(* IEC 61131-3 sources: plc-process-lib/tests/POUs/Suites/FB_Util_Test, 29 files *)

(* ---- IsFiniteAboveSaneMaxReturnsFalse.method.decl.st ---- *)
// F_IsFinite: |x| > REAL_SANE_MAX — мусор (перепутан порядок слов Modbus): 1e31, -1e31 и
// наибольшее REAL — FALSE.
METHOD PRIVATE IsFiniteAboveSaneMaxReturnsFalse
VAR
    uBits : U_RealBits;      // значение REAL по битам IEEE 754
END_VAR

(* ---- IsFiniteInfReturnsFalse.method.decl.st ---- *)
// F_IsFinite: +Inf и -Inf — FALSE.
METHOD PRIVATE IsFiniteInfReturnsFalse
VAR
    uBits : U_RealBits;      // значение REAL по битам IEEE 754
END_VAR

(* ---- IsFiniteNaNReturnsFalse.method.decl.st ---- *)
// F_IsFinite: тихий NaN с обоими знаками и с полной мантиссой — FALSE (проверка R4 контракта).
METHOD PRIVATE IsFiniteNaNReturnsFalse
VAR
    uBits : U_RealBits;      // значение REAL по битам IEEE 754
END_VAR

(* ---- IsFiniteNormalReturnsTrue.method.decl.st ---- *)
// F_IsFinite: обычные числа, 0, -0, наименьшее денормализованное и граница ±REAL_SANE_MAX
// (включительно) — TRUE.
METHOD PRIVATE IsFiniteNormalReturnsTrue
VAR
    uBits : U_RealBits;      // значение REAL по битам IEEE 754
END_VAR

(* ---- LimitMonitorDisabledNeverSets.method.decl.st ---- *)
// Выключенная уставка (xEnable = FALSE) не взводит флаг: 10 с значение далеко за уставкой.
METHOD PRIVATE LimitMonitorDisabledNeverSets
VAR
    fbTime   : FB_FakeTime;       // подменное время
    fbLim    : FB_LimitMonitor;   // ФБ под тестом
    stLimCfg : ST_AiLimitCfg;     // параметры уставки
    iStep : INT;             // шаг цикла
    xEverSet : BOOL;            // флаг взводился хотя бы раз
END_VAR

(* ---- LimitMonitorDisabledNeverSets.method.impl.st ---- *)
coUnit.TEST('Util_LimitMonitor_Disabled_NeverSets');

stLimCfg.xEnable := FALSE;
stLimCfg.rSetpoint_eu := 50.0;
FOR iStep := 1 TO 100 DO
    fbTime.Advance(tStep := T#100MS);
    fbLim(rValue_eu := 90.0, xHighLimit := TRUE, stCfg := stLimCfg, itfTime := fbTime);
    xEverSet := xEverSet OR fbLim.xOut OR fbLim.xRaw;
END_FOR
AssertFalse(Condition := xEverSet, Message := 'disabled limit must never set the flag');

coUnit.TEST_FINISHED();

(* ---- LimitMonitorForceOffClearsImmediately.method.decl.st ---- *)
// xForceOff снимает флаг и сырой флаг в том же вызове, несмотря на задержку снятия 10 с; после
// снятия xForceOff флаг возвращается (значение по-прежнему выше уставки, задержки включения нет).
METHOD PRIVATE LimitMonitorForceOffClearsImmediately
VAR
    fbTime   : FB_FakeTime;       // подменное время
    fbLim    : FB_LimitMonitor;   // ФБ под тестом
    stLimCfg : ST_AiLimitCfg;     // параметры уставки
END_VAR

(* ---- LimitMonitorHighHysteresisClearsBelowSpMinusHyst.method.decl.st ---- *)
// Верхняя уставка 80, гистерезис 5: флаг при значении >= 80 (включительно), держится до 75
// включительно, снимается ниже 75; в зоне гистерезиса снятый флаг не возвращается.
METHOD PRIVATE LimitMonitorHighHysteresisClearsBelowSpMinusHyst
VAR
    fbTime   : FB_FakeTime;       // подменное время
    fbLim    : FB_LimitMonitor;   // ФБ под тестом
    stLimCfg : ST_AiLimitCfg;     // параметры уставки
END_VAR

(* ---- LimitMonitorLowHysteresisClearsAboveSpPlusHyst.method.decl.st ---- *)
// Нижняя уставка 20, гистерезис 2 — зеркально: флаг при значении <= 20, держится до 22
// включительно, снимается выше 22.
METHOD PRIVATE LimitMonitorLowHysteresisClearsAboveSpPlusHyst
VAR
    fbTime   : FB_FakeTime;       // подменное время
    fbLim    : FB_LimitMonitor;   // ФБ под тестом
    stLimCfg : ST_AiLimitCfg;     // параметры уставки
END_VAR

(* ---- LimitMonitorNonFiniteValueKeepsState.method.decl.st ---- *)
// Неконечное значение (NaN, ±Inf, больше REAL_SANE_MAX) флаг не меняет: -Inf не снимает
// взведённый флаг верхней уставки, +Inf не взводит снятый.
METHOD PRIVATE LimitMonitorNonFiniteValueKeepsState
VAR
    fbTime   : FB_FakeTime;       // подменное время
    fbLim    : FB_LimitMonitor;   // ФБ под тестом
    stLimCfg : ST_AiLimitCfg;     // параметры уставки
    uBits : U_RealBits;      // значение REAL по битам IEEE 754
END_VAR

(* ---- LimitMonitorOffDelayHoldsFlag.method.decl.st ---- *)
// Задержка снятия 2 с: сырой флаг снимается сразу, выходной держится до t0 + 1,9 с и снимается
// ровно в t0 + 2,0 с.
METHOD PRIVATE LimitMonitorOffDelayHoldsFlag
VAR
    fbTime   : FB_FakeTime;       // подменное время
    fbLim    : FB_LimitMonitor;   // ФБ под тестом
    stLimCfg : ST_AiLimitCfg;     // параметры уставки
    iStep : INT;             // шаг цикла
END_VAR

(* ---- LimitMonitorOffDelayHoldsFlag.method.impl.st ---- *)
coUnit.TEST('Util_LimitMonitor_OffDelay_HoldsFlag');

stLimCfg.xEnable := TRUE;
stLimCfg.rSetpoint_eu := 80.0;
stLimCfg.rHyst_eu := 2.0;
stLimCfg.tOffDelay := T#2S;
fbLim(rValue_eu := 85.0, xHighLimit := TRUE, stCfg := stLimCfg, itfTime := fbTime);
AssertTrue(Condition := fbLim.xOut, Message := 'flag set without on-delay');
fbLim(rValue_eu := 70.0, xHighLimit := TRUE, stCfg := stLimCfg, itfTime := fbTime);    // t0
AssertFalse(Condition := fbLim.xRaw, Message := 'raw flag cleared at once');
FOR iStep := 1 TO 19 DO
    fbTime.Advance(tStep := T#100MS);
    fbLim(rValue_eu := 70.0, xHighLimit := TRUE, stCfg := stLimCfg, itfTime := fbTime);
END_FOR
AssertTrue(Condition := fbLim.xOut, Message := 'flag held at t0 + 1.9 s');
fbTime.Advance(tStep := T#100MS);
fbLim(rValue_eu := 70.0, xHighLimit := TRUE, stCfg := stLimCfg, itfTime := fbTime);
AssertFalse(Condition := fbLim.xOut, Message := 'flag cleared exactly at t0 + 2.0 s');

coUnit.TEST_FINISHED();

(* ---- LimitMonitorOnDelayShortExcursionIgnored.method.decl.st ---- *)
// Задержка срабатывания 3 с: выброс 2,9 с за уставку флаг не взводит (сырой флаг — да);
// устойчивое превышение — флаг ровно через 3 с.
METHOD PRIVATE LimitMonitorOnDelayShortExcursionIgnored
VAR
    fbTime   : FB_FakeTime;       // подменное время
    fbLim    : FB_LimitMonitor;   // ФБ под тестом
    stLimCfg : ST_AiLimitCfg;     // параметры уставки
    iStep : INT;             // шаг цикла
    xEverSet : BOOL;            // флаг взводился хотя бы раз
END_VAR

(* ---- LimitMonitorOnDelayShortExcursionIgnored.method.impl.st ---- *)
coUnit.TEST('Util_LimitMonitor_OnDelay_ShortExcursionIgnored');

stLimCfg.xEnable := TRUE;
stLimCfg.rSetpoint_eu := 80.0;
stLimCfg.rHyst_eu := 2.0;
stLimCfg.tOnDelay := T#3S;
fbLim(rValue_eu := 85.0, xHighLimit := TRUE, stCfg := stLimCfg, itfTime := fbTime);    // t0
FOR iStep := 1 TO 29 DO                                                               // t0 + 2,9 с
    fbTime.Advance(tStep := T#100MS);
    fbLim(rValue_eu := 85.0, xHighLimit := TRUE, stCfg := stLimCfg, itfTime := fbTime);
    xEverSet := xEverSet OR fbLim.xOut;
END_FOR
AssertTrue(Condition := fbLim.xRaw, Message := 'raw flag is set before the delay');
fbTime.Advance(tStep := T#100MS);
fbLim(rValue_eu := 70.0, xHighLimit := TRUE, stCfg := stLimCfg, itfTime := fbTime);    // t0 + 3,0 с
xEverSet := xEverSet OR fbLim.xOut;
AssertFalse(Condition := xEverSet, Message := 'excursion shorter than the on-delay must be ignored');
fbLim(rValue_eu := 85.0, xHighLimit := TRUE, stCfg := stLimCfg, itfTime := fbTime);    // t1
FOR iStep := 1 TO 29 DO
    fbTime.Advance(tStep := T#100MS);
    fbLim(rValue_eu := 85.0, xHighLimit := TRUE, stCfg := stLimCfg, itfTime := fbTime);
END_FOR
AssertFalse(Condition := fbLim.xOut, Message := 'no flag at t1 + 2.9 s');
fbTime.Advance(tStep := T#100MS);
fbLim(rValue_eu := 85.0, xHighLimit := TRUE, stCfg := stLimCfg, itfTime := fbTime);    // t1 + 3,0 с
AssertTrue(Condition := fbLim.xOut, Message := 'flag exactly at t1 + 3.0 s');

coUnit.TEST_FINISHED();

(* ---- LimitMonitorReenabledRestartsOnDelay.method.decl.st ---- *)
// Выключение уставки во время задержки срабатывания (2 с) сбрасывает отсчёт: после повторного
// включения в t0 + 1,6 с флаг — ровно через 2 с от включения, а не в t0 + 2,0 с.
METHOD PRIVATE LimitMonitorReenabledRestartsOnDelay
VAR
    fbTime   : FB_FakeTime;       // подменное время
    fbLim    : FB_LimitMonitor;   // ФБ под тестом
    stLimCfg : ST_AiLimitCfg;     // параметры уставки
    iStep : INT;             // шаг цикла
END_VAR

(* ---- LimitMonitorReenabledRestartsOnDelay.method.impl.st ---- *)
coUnit.TEST('Util_LimitMonitor_Reenabled_RestartsOnDelay');

stLimCfg.xEnable := TRUE;
stLimCfg.rSetpoint_eu := 80.0;
stLimCfg.tOnDelay := T#2S;
fbLim(rValue_eu := 90.0, xHighLimit := TRUE, stCfg := stLimCfg, itfTime := fbTime);    // t0
FOR iStep := 1 TO 15 DO                                                               // t0 + 1,5 с
    fbTime.Advance(tStep := T#100MS);
    fbLim(rValue_eu := 90.0, xHighLimit := TRUE, stCfg := stLimCfg, itfTime := fbTime);
END_FOR
stLimCfg.xEnable := FALSE;
fbLim(rValue_eu := 90.0, xHighLimit := TRUE, stCfg := stLimCfg, itfTime := fbTime);
AssertFalse(Condition := fbLim.xOut OR fbLim.xRaw, Message := 'disabled: flags cleared');
stLimCfg.xEnable := TRUE;
FOR iStep := 1 TO 5 DO                                                                // t0 + 1,6 … 2,0 с
    fbTime.Advance(tStep := T#100MS);
    fbLim(rValue_eu := 90.0, xHighLimit := TRUE, stCfg := stLimCfg, itfTime := fbTime);
END_FOR
AssertFalse(Condition := fbLim.xOut, Message := 'old timing must not complete after re-enable');
FOR iStep := 1 TO 15 DO                                                               // t0 + 3,5 с
    fbTime.Advance(tStep := T#100MS);
    fbLim(rValue_eu := 90.0, xHighLimit := TRUE, stCfg := stLimCfg, itfTime := fbTime);
END_FOR
AssertFalse(Condition := fbLim.xOut, Message := 'no flag 1.9 s after re-enable');
fbTime.Advance(tStep := T#100MS);
fbLim(rValue_eu := 90.0, xHighLimit := TRUE, stCfg := stLimCfg, itfTime := fbTime);    // t0 + 3,6 с
AssertTrue(Condition := fbLim.xOut, Message := 'flag 2.0 s after re-enable');

coUnit.TEST_FINISHED();

(* ---- RateLimitLrNonFiniteTargetOrZeroDtHoldsCurrent.method.decl.st ---- *)
// F_RateLimitLr: цель NaN (мусор Modbus) или шаг времени 0 — значение не меняется; скорость 0 — сразу к цели;
// текущее значение NaN — сразу к цели (как F_RateLimit, F-11).
METHOD PRIVATE RateLimitLrNonFiniteTargetOrZeroDtHoldsCurrent
VAR
    uBits : U_RealBits;      // значение REAL по битам IEEE 754
    lrOut : LREAL;           // результат F_RateLimitLr
    lrNaN : LREAL;           // NaN в LREAL
END_VAR

(* ---- RateLimitLrSmallStepNotLost.method.decl.st ---- *)
// F_RateLimitLr: состояние в LREAL — 1000 шагов по 1 мс со скоростью 0,003 ед./с от 70,0 дают 70,003 (в REAL
// приращение 3·10⁻⁶ меньше половины шага REAL рядом с 70 и терялось бы); спад — так же; цель достигается точно.
METHOD PRIVATE RateLimitLrSmallStepNotLost
VAR
    lrUp   : LREAL;          // рост: состояние рампы
    lrDown : LREAL;          // спад: состояние рампы
    iStep  : INT;            // шаг цикла
END_VAR

(* ---- RateLimitLrSmallStepNotLost.method.impl.st ---- *)
coUnit.TEST('Util_RateLimitLr_SmallStep_NotLost');

lrUp := 70.0;
lrDown := 70.0;
FOR iStep := 1 TO 1000 DO
    lrUp := F_RateLimitLr(lrCurrent := lrUp, rTarget := 100.0, rRateUp_ups := 0.003, rRateDown_ups := 0.003,
                          lrDt_s := 0.001);
    lrDown := F_RateLimitLr(lrCurrent := lrDown, rTarget := 0.0, rRateUp_ups := 0.003, rRateDown_ups := 0.003,
                            lrDt_s := 0.001);
END_FOR
// ожидаемое: 70 ± 0,003 · 1 с; допуск — шаг REAL скорости 0,003 · 1000 шагов
AssertEquals_LREAL(Expected := LREAL#70.003, Actual := lrUp, Delta := LREAL#1.0E-7, Message := 'ramp up not lost');
AssertEquals_LREAL(Expected := LREAL#69.997, Actual := lrDown, Delta := LREAL#1.0E-7, Message := 'ramp down not lost');
AssertEquals_LREAL(Expected := LREAL#42.5, Actual := F_RateLimitLr(lrCurrent := LREAL#42.49, rTarget := 42.5,
                   rRateUp_ups := 1.0, rRateDown_ups := 1.0, lrDt_s := 1.0), Delta := LREAL#0.0,
                   Message := 'reaches the target exactly');

coUnit.TEST_FINISHED();

(* ---- RateLimitNonFiniteCurrentJumpsToTarget.method.decl.st ---- *)
// F_RateLimit: текущее значение NaN (мусор прошлого шага) заменяется конечной целью — ограничитель
// не застревает на NaN.
METHOD PRIVATE RateLimitNonFiniteCurrentJumpsToTarget
VAR
    uBits : U_RealBits;      // значение REAL по битам IEEE 754
    rOut  : REAL;            // результат F_RateLimit
END_VAR

(* ---- RateLimitNonFiniteTargetHoldsCurrent.method.decl.st ---- *)
// F_RateLimit: цель NaN, +Inf или больше REAL_SANE_MAX (мусор из Modbus/ПИД) — значение удерживается.
METHOD PRIVATE RateLimitNonFiniteTargetHoldsCurrent
VAR
    uBits : U_RealBits;      // значение REAL по битам IEEE 754
    rOut  : REAL;            // результат F_RateLimit
END_VAR

(* ---- StartsWindowClearEmpties.method.decl.st ---- *)
// Clear очищает окно: пусков 0, освобождать нечего.
METHOD PRIVATE StartsWindowClearEmpties
VAR
    fbWin : FB_StartsWindow; // ФБ под тестом
END_VAR

(* ---- StartsWindowCountsOnlyLastHour.method.decl.st ---- *)
// FB_StartsWindow: пуски в 1:00, 1:20, 1:40 — в окне последнего часа их 3, 2, 1, 0 по мере
// старения. Источник: tools/reference/common.py, сценарий starts_window.
METHOD PRIVATE StartsWindowCountsOnlyLastHour
VAR
    fbWin : FB_StartsWindow; // ФБ под тестом
END_VAR

(* ---- StartsWindowExactlyOneHourOldNotCounted.method.decl.st ---- *)
// Граница окна: отметка ровно часовой давности уже не считается (ltNow - t < STARTS_WINDOW).
METHOD PRIVATE StartsWindowExactlyOneHourOldNotCounted
VAR
    fbWin : FB_StartsWindow; // ФБ под тестом
END_VAR

(* ---- StartsWindowRingCapacityMatchesConst.method.decl.st ---- *)
// Ёмкость кольца altStart равна GVL_Const.STARTS_WINDOW_MAX: индексы кольца считаются по константе,
// тест ловит расхождение, если границу массива запишут числом.
// Тест обращается к внутренней переменной ФБ намеренно: это проверка раскладки, а не API.
METHOD PRIVATE StartsWindowRingCapacityMatchesConst
VAR
    fbWin : FB_StartsWindow; // ФБ под тестом
    ltOne : LTIME;           // один элемент кольца
END_VAR

(* ---- StartsWindowRingFullOverwritesOldest.method.decl.st ---- *)
// Кольцо на STARTS_WINDOW_MAX = 30: 31 пуск с шагом 1 мин (1:00…1:30) — остаются 30 последних;
// в 1:30 при лимите 30 окно освободится через 31 мин (самый старый оставшийся — 1:01).
// Источник: tools/reference/common.py, сценарий starts_window.
METHOD PRIVATE StartsWindowRingFullOverwritesOldest
VAR
    fbWin : FB_StartsWindow; // ФБ под тестом
    ltStart : LTIME := LTIME#1H;   // время очередного пуска
    iStep : INT;             // шаг цикла
END_VAR

(* ---- StartsWindowRingFullOverwritesOldest.method.impl.st ---- *)
coUnit.TEST('Util_StartsWindow_RingFull_OverwritesOldest');

FOR iStep := 0 TO 30 DO
    fbWin.Register(ltNow := ltStart);
    ltStart := ltStart + LTIME#1M;
END_FOR
AssertEquals_UINT(Expected := 30, Actual := fbWin.Count(ltNow := LTIME#1H30M), Message := 'ring keeps 30 starts');
AssertEquals_LTIME(Expected := LTIME#31M, Actual := fbWin.TimeToFree(ltNow := LTIME#1H30M, uiMax := 30),
                   Message := 'the start of 1:00 was overwritten, the oldest kept is 1:01');

coUnit.TEST_FINISHED();

(* ---- StartsWindowTimeBackwardsDropsFutureStamps.method.decl.st ---- *)
// Время назад: отметки «из будущего» удаляются и в Count, и в Register; окно остаётся упорядоченным.
METHOD PRIVATE StartsWindowTimeBackwardsDropsFutureStamps
VAR
    fbWin : FB_StartsWindow; // ФБ под тестом
END_VAR

(* ---- StartsWindowTimeToFreeReportsRemaining.method.decl.st ---- *)
// TimeToFree: пуски 1:00, 1:10, 1:20; в 1:30 при лимите 3 — 30 мин, при лимите 2 — 40 мин,
// при лимите 4 и без лимита (0) — 0; в 2:00 при лимите 3 — 0.
// Источник: tools/reference/common.py, сценарий starts_window.
METHOD PRIVATE StartsWindowTimeToFreeReportsRemaining
VAR
    fbWin : FB_StartsWindow; // ФБ под тестом
END_VAR
